Fanuc KAREL source: kb00069.KL

-- PROVISIONAL review KL for V1013-1; original PC SHA256 f811c0cc2fcf43d5b22f7808c0e405813b6dc56712a767c5be51f4c92934e9a7
-- Incomplete behavior may be omitted. Consult companion uncertainty JSON. Do not deploy.
PROGRAM KB00069
%NOLOCKGROUP
BEGIN
  -- UNRESOLVED_PC offsets 5-14; opcodes 3F,75
  -- UNRESOLVED_PC offsets 19-26; opcodes 9D,23
  -- UNRESOLVED_PC offsets 31-40; opcodes 3F,75
  -- UNRESOLVED_PC offsets 45-52; opcodes 9D,23
  -- UNRESOLVED_PC offsets 57-89; opcodes 27,22,2A,22,22,2A,22,31
  -- UNRESOLVED_PC offsets 94-98; opcodes 7F
END KB00069
